(* IEC 61131-3 sources: structured-text/samples/unsupported/string, 2 files *)

(* ---- t17-5.st ---- *)
PROGRAM Test
	VAR
		CONDITION_RED : BOOL;
		IBOUNCE : WORD ;
		MYDUB : DWORD ;
		AWORD, BWORD, CWORD : INT;
		MYSTR: STRING[10] ;
	END_VAR
END_PROGRAM

(* ---- t18-5.st ---- *)
PROGRAM Test
	VAR
  		MYBIT : BOOL := 1 ;
  		OKAY : STRING[10] := 'OK';
	END_VAR
END_PROGRAM
